Universal Robots URScript: T014_qwen2.5-coder_32b_baseline_rep1.urscript

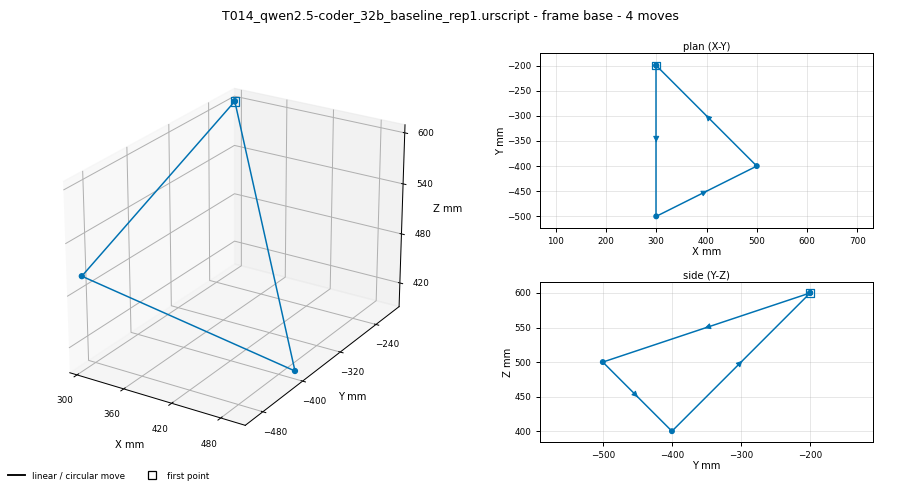
[picture p0: tool path of T014_qwen2.5-coder_32b_baseline_rep1.urscript in frame base, 4 of 6 moves have a stored position in this frame; points joined in program order, loops and branches not executed]
def hybrid_multi_angle_inspection():
    # Move to Home position
    movej(get_inverse_kin([0, -90, 90, -90, 45, 0]), a=1.2, v=1.05)

    # Move to Top-down view position
    movel(p[0.3, -0.2, 0.6, 3.14159, 0, 0], a=1.2, v=0.75)

    # Move to Side view position
    movel(p[0.3, -0.5, 0.5, 3.14159, 0, 1.57], a=1.2, v=0.6)

    # Move to Angled view position
    movel(p[0.5, -0.4, 0.4, 3.14159, 0, 1.0], a=1.2, v=0.6)

    # Retract
    movel(p[0.3, -0.2, 0.6, 3.14159, 0, 0], a=1.2, v=0.75)

    # Move back to Home position
    movej(get_inverse_kin([0, -90, 90, -90, 45, 0]), a=1.2, v=1.05)
end

hybrid_multi_angle_inspection()
